FUNCTION_BLOCK RUL_ESTIMATION
  {SET_ATTRIBUTE(OpcUa, SERVICE)}
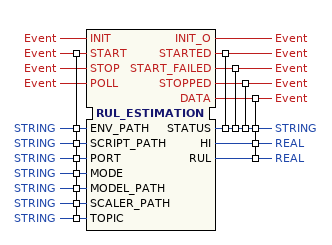
  EVENT_INPUT
    INIT;
    START WITH ENV_PATH, SCRIPT_PATH, PORT, MODE, MODEL_PATH, SCALER_PATH, TOPIC;
    STOP;
    POLL;
  END_EVENT
  EVENT_OUTPUT
    INIT_O;
    STARTED WITH STATUS;
    START_FAILED WITH STATUS;
    STOPPED WITH STATUS;
    DATA WITH HI, RUL, STATUS;
  END_EVENT
  VAR_INPUT
    ENV_PATH : STRING; {SET_ATTRIBUTE(OpcUa, Variable)}
    SCRIPT_PATH : STRING; {SET_ATTRIBUTE(OpcUa, Variable)}
    PORT : STRING; {SET_ATTRIBUTE(OpcUa, Variable)}
    MODE : STRING; {SET_ATTRIBUTE(OpcUa, Variable)}
    MODEL_PATH : STRING; {SET_ATTRIBUTE(OpcUa, Variable)}
    SCALER_PATH : STRING; {SET_ATTRIBUTE(OpcUa, Variable)}
    TOPIC : STRING; {SET_ATTRIBUTE(OpcUa, Variable)}
  END_VAR
  VAR_OUTPUT
    STATUS : STRING; {SET_ATTRIBUTE(OpcUa, Variable)}
    HI : REAL; {SET_ATTRIBUTE(OpcUa, Variable)}
    RUL : REAL; (* Remaining useful life in hours (-1 = no estimate yet) *) {SET_ATTRIBUTE(OpcUa, Variable)}
  END_VAR
END_FUNCTION_BLOCK
